PROGRAM Gr01Control
VAR_INPUT
	(* Input variables / Eingang Variablen *)
	bEnable						:BOOL;						(* Enable Gr01Control *)

	(* Instances *)
	fbAxisSawBow				:FB_Gr01SawBow;
	fbAxisAngle					:FB_Gr01Angle;

	fbSawband			 		:FB_Gr01Sawband;

END_VAR
VAR
	(* Enummerations *)

	(* Variables *)
	bAllAxisCtrlEnabled				:BOOL;						(* All axis have controller enabled *)
	bAllAxisStandStill				:BOOL;						(* All axis stand still *)
	bAllAxisNotMoving				:BOOL;						(* All axis not moving *)
	bAllAxisReferenced				:BOOL;						(* All axis referenced *)
	
	BandDistance_m					:LREAL;
	rMachineSawbandSpeed_mmin		:LREAL;

	(* References *)

	(* Interfaces *)

	(* Instances *)
	fbAlarm						:FB_Gr01Alarm;
	fbSafety					:FB_Gr01Safety;
	fbSignals					:FB_Gr01Signals;
	fbUtility					:FB_Gr01Utility;
	rtBtnStart					:R_TRIG;
	
	SawbandVelo					:FB_PosVeloEnc;
	fbLowPassFilter				:FB_LowPassFilter;
	tonSawBandVeloErr			:TON;
	tonSawBandInVelo			:TON;
	TimerVelo					:TON;

END_VAR
VAR CONSTANT
	nFatalErrorMaxIdx			:INT := 0;						(* Maximal index of  using alarms *)
	nErrorMaxIdx				:INT := 19;					(* Maximal index of  using alarms *)
	nWarningMaxIdx				:INT := 0;						(* Maximal index of  using alarms *)
	nMessageMaxIdx				:INT := 1;						(* Maximal index of  using alarms *)
	nHintMaxIdx					:INT := 0;						(* Maximal index of  using alarms *)

	dnFatalErrorBaseIdentNo		:DINT := 11000;				(* Fatal error identification number *)
	dnErrorBaseIdentNo			:DINT := 11100;				(* Error identification number *)
	dnWarningBaseIdentNo		:DINT := 11200;				(* Warning identification number *)
	dnMessageBaseIdentNo		:DINT := 11300;				(* Message identification number *)
	dnHintBaseIdentNo			:DINT := 11400;				(* Hint identification number *)
END_VAR

IF NOT bEnable
THEN
	RETURN;
END_IF;

A_Utility();
A_Safety();
A_Axis();
A_Sawband();
A_Signals();
A_Alarm();

ACTION A_Alarm:

(* Collect and execute input alarms *)
fbAlarm.stAlarmIn.arbError[0].bActive := NOT binGr01LightCurtainOK
                                                		      AND (Gr01Home.fbProcedure.bBusy
                                                      				OR Gr01Auto.fbProcedure.bBusy);
fbAlarm.stAlarmIn.arbError[0].dnCode := dnErrorBaseIdentNo + 0;

fbAlarm.stAlarmIn.arbError[1].bActive := NOT binGr01SawbandRelease
								    AND bgGr00ModeAutomatic
								    AND bgGr00MachineRunning;
fbAlarm.stAlarmIn.arbError[1].dnCode := dnErrorBaseIdentNo + 1;

fbAlarm.stAlarmIn.arbError[2].bActive := FALSE;
fbAlarm.stAlarmIn.arbError[2].dnCode := dnErrorBaseIdentNo + 2;

fbAlarm.stAlarmIn.arbError[3].bActive := FALSE;
fbAlarm.stAlarmIn.arbError[3].dnCode := dnErrorBaseIdentNo + 3;

fbAlarm.stAlarmIn.arbError[4].bActive := fbAxisSawBow.bErrorTerminal;
fbAlarm.stAlarmIn.arbError[4].dnCode := dnErrorBaseIdentNo + 4;

fbAlarm.stAlarmIn.arbError[5].bActive := fbAxisSawBow.fbController.bErrorInit;
fbAlarm.stAlarmIn.arbError[5].dnCode := dnErrorBaseIdentNo + 5;

fbAlarm.stAlarmIn.arbError[6].bActive := fbAxisSawBow.bErrorCtrlEnabled;
fbAlarm.stAlarmIn.arbError[6].dnCode := dnErrorBaseIdentNo + 6;

fbAlarm.stAlarmIn.arbError[7].bActive := fbAxisSawBow.fbController.bError OR fbAxisSawBow.fbMoveManual.bError OR fbAxisSawBow.fbMoveAuto.bError;
fbAlarm.stAlarmIn.arbError[7].dnCode := dnErrorBaseIdentNo + 7;

fbAlarm.stAlarmIn.arbError[8].bActive := fbAxisAngle.bErrorTerminal;
fbAlarm.stAlarmIn.arbError[8].dnCode := dnErrorBaseIdentNo + 8;

fbAlarm.stAlarmIn.arbError[9].bActive := fbAxisAngle.fbController.bErrorInit;
fbAlarm.stAlarmIn.arbError[9].dnCode := dnErrorBaseIdentNo + 9;

fbAlarm.stAlarmIn.arbError[10].bActive := fbAxisAngle.bErrorCtrlEnabled;
fbAlarm.stAlarmIn.arbError[10].dnCode := dnErrorBaseIdentNo + 10;

fbAlarm.stAlarmIn.arbError[11].bActive := fbAxisAngle.fbController.bError OR fbAxisAngle.fbMoveManual.bError OR fbAxisAngle.fbMoveAuto.bError;
fbAlarm.stAlarmIn.arbError[11].dnCode := dnErrorBaseIdentNo + 11;

fbAlarm.stAlarmIn.arbError[12].bActive := fbSawband.bErrorTerminal;
fbAlarm.stAlarmIn.arbError[12].dnCode := dnErrorBaseIdentNo + 12;

fbAlarm.stAlarmIn.arbError[13].bActive := fbSawband.fbController.bErrorInit;
fbAlarm.stAlarmIn.arbError[13].dnCode := dnErrorBaseIdentNo + 13;

fbAlarm.stAlarmIn.arbError[14].bActive := fbSawband.bErrorCtrlEnabled;
fbAlarm.stAlarmIn.arbError[14].dnCode := dnErrorBaseIdentNo + 14;

fbAlarm.stAlarmIn.arbError[15].bActive := fbSawband.fbController.bError OR fbSawband.fbMoveManual.bError OR fbSawband.fbMoveAuto.bError;
fbAlarm.stAlarmIn.arbError[15].dnCode := dnErrorBaseIdentNo + 15;

fbAlarm.stAlarmIn.arbError[16].bActive := FALSE;
fbAlarm.stAlarmIn.arbError[16].dnCode := dnErrorBaseIdentNo + 16;

fbAlarm.stAlarmIn.arbError[17].bActive := GVL_Gr0100.bgGr01SawbandVeloError_1;
fbAlarm.stAlarmIn.arbError[17].dnCode := dnErrorBaseIdentNo + 17;

fbAlarm.stAlarmIn.arbError[18].bActive := GVL_Gr0100.bgGr01SawbandVeloError_2;
fbAlarm.stAlarmIn.arbError[18].dnCode := dnErrorBaseIdentNo + 18;

fbAlarm.stAlarmIn.arbError[19].bActive := (* bgGr00MachineRunning
							AND fbSawband.bCtrlEnabled
							AND fbSawband.bSpeedReached
							AND *) NOT fbSafety.bPipeNotInCrashArea;  (* 20260219 ES/KG *)

fbAlarm.stAlarmIn.arbError[19].dnCode := dnErrorBaseIdentNo + 19;

fbAlarm.stAlarmIn.arbWarning[0].bActive := fbSawband.bErrorVacuumCleanerNOK;
fbAlarm.stAlarmIn.arbWarning[0].dnCode := dnWarningBaseIdentNo + 0;

fbAlarm.stAlarmIn.arbMessage[0].bActive := NOT binGr01LightCurtainOK
							      AND NOT fbAlarm.stAlarmIn.arbError[0].bActive
							      AND NOT fbAlarm.stAlarmOut.arbError[0].bActive;
fbAlarm.stAlarmIn.arbMessage[0].dnCode := dnMessageBaseIdentNo + 0;

fbAlarm.stAlarmIn.arbMessage[1].bActive := NOT binGr01SawbandRelease;
fbAlarm.stAlarmIn.arbMessage[1].dnCode := dnMessageBaseIdentNo + 1;

(* Execute utility *)
fbAlarm(
	etMachineMode := etgGr00MachineMode,
	etMachineState := etgGr00MachineState,
	bNoEStop := bgGr00NoEmergencyStop,
	bConfirmAlarm := bgGr00ConfirmAlarm,
	dtDateTime := stgGr00DateTime.dtDateTime,
	nFatalErrorMaxIdx := nFatalErrorMaxIdx,
	nErrorMaxIdx := nErrorMaxIdx,
	nWarningMaxIdx := nWarningMaxIdx,
	nMessageMaxIdx := nMessageMaxIdx,
	nHintMaxIdx := nHintMaxIdx,
	bMoveInterrupted := bgGr01MoveInterrupted,
	bHomeCompleted := bgGr01HomeCompleted,
	stAlarmOut => stgGr01Alarm.stControl
);
END_ACTION

ACTION A_Axis:

(* Enable axis saw bow *)
stgGr01HMI.stHMITOPLC.lrAxisSawBowNoRefVelo := 10;

fbAxisSawBow(
	bEnable						:= TRUE,
	etMachineMode				:= etgGr00MachineMode,
	etMachineState				:= etgGr00MachineState,
	bMachineStandstill			:= bgGr00MachineStandstill,
	bNoEStop					:= bgGr00NoEmergencyStop,
	bPowerSupplyOn				:= bgGr00PowerSupplyOk,
	bSafetyOK					:= bgGr01LightCurtainOK
								   AND bgGr00AllDoorsClosedLocked,
	bCtrlInterrupt				:= FALSE,
	bMoveRelease				:= TRUE,
	bPlusRelease				:= TRUE,
	bMinusRelease				:= TRUE,
	bSignalReference			:= NOT binGr01AxisSawBowLimitMax,
	bSignalHWLimitMax			:= NOT binGr01AxisSawBowLimitMax,
	bSignalHWLimitMin			:= NOT binGr01AxisSawBowLimitMin,
	lrSoftLimitMax				:= stgGr01HMI.stHMITOPLC.lrAxisSawBowSoftLimitMax,
	lrSoftLimitMin				:= stgGr01HMI.stHMITOPLC.lrAxisSawBowSoftLimitMin,
	bConfirmAlarm				:= bgGr00ConfirmAlarm,
	bTipPlus					:= stgGr01HMI.stHMITOPLC.bBtnAxisSawBowPlus,
	bTipMinus					:= stgGr01HMI.stHMITOPLC.bBtnAxisSawBowMinus,
	lrManualVelocity			:= stgGr01HMI.stHMITOPLC.lrAxisSawBowManualVelo,
	lrNoRefVelocity				:= stgGr01HMI.stHMITOPLC.lrAxisSawBowNoRefVelo,
	bVelocityLimitEn			:= FALSE,
	lrAcceleration				:= 100.0,
	lrDeceleration				:= 100.0,
	lrJerk						:= 100.0,
	lrOverride					:= fbUtility.rActOverride,
	lrExtOverride				:= 0.0,
	dnRatioNumerator			:= 1,
	udnRatioDenominator			:= 1,
	bEngineTorqueLimitEn		:= FALSE,
	lrEngineTorque				:= 200.0,
	tControllerOff				:= tgGr01ControllerOff,
	bWithAbsoluteEncoder		:= FALSE,
	lrOriginShiftPos			:= stgGr01HMI.stHMITOPLC.lrAxisSawBowOriginShiftPos,
	bVeloForceCtrlEn			:= FALSE,
	tAdsTimeOut					:= DEFAULT_ADS_TIMEOUT,
	bHomeCompleted				:= bgGr01HomeCompleted,
	Drive						:= GVL_Gr01Interface.igGr01DriveSawBow,
	Axis						:= GVL_Gr01Interface.igGr01AxisSawBow,
	MasterAxis					:= GVL_Gr00Interface.iAxisDummy,
	
	lrActPosition				=> stgGr01HMI.stPLCTOHMI.lrAxisSawBowActPos,
	lrActVelocity				=> stgGr01HMI.stPLCTOHMI.lrAxisSawBowActVelo,
	lrActForce					=> stgGr01HMI.stPLCTOHMI.lrAxisSawBowActForce
);

(* Enable Axis angle *)
stgGr01HMI.stHMITOPLC.lrAxisAngleNoRefVelo := 10;



fbAxisAngle(
	bEnable						:= TRUE,

	etMachineMode				:= etgGr00MachineMode,
	etMachineState				:= etgGr00MachineState,
	bMachineStandstill			:= bgGr00MachineStandstill,
	bNoEStop					:= bgGr00NoEmergencyStop,
	bPowerSupplyOn				:= bgGr00PowerSupplyOk,
	bSafetyOK					:= bgGr01LightCurtainOK
								   AND bgGr00AllDoorsClosedLocked,
	bCtrlInterrupt				:= FALSE,
	bMoveRelease				:= TRUE,
	bMoveInterrupt				:= FALSE,
	bPlusRelease				:= TRUE,
	bMinusRelease				:= TRUE,	(*stgGr00HMI.stHMITOPLC.bSafetyInterlockOff*)
	bHWSignalLimitMax			:= NOT binGr01AxisAngleLimitMax,
	bHWSignalLimitMin			:= NOT binGr01AxisAngleLimitMin,
	lrSoftLimitMax				:= stgGr01HMI.stHMITOPLC.lrAxisAngleSoftLimitMax,
	lrSoftLimitMin				:= stgGr01HMI.stHMITOPLC.lrAxisAngleSoftLimitMin,
	bConfirmAlarm				:= bgGr00ConfirmAlarm,
	bTipPlus					:= stgGr01HMI.stHMITOPLC.bBtnAxisAnglePlus,
	bTipMinus					:= stgGr01HMI.stHMITOPLC.bBtnAxisAngleMinus,
	lrManualVelocity			:= stgGr01HMI.stHMITOPLC.lrAxisAngleManualVelo,
	lrVelocityNoRef				:= stgGr01HMI.stHMITOPLC.lrAxisAngleNoRefVelo,
	bVelocityLimitEn			:= FALSE,
	lrAcceleration				:= 100.0,
	lrDeceleration				:= 100.0,
	lrJerk						:= 100.0,
	lrOverride					:= fbUtility.rActOverride,
	bEngineTorqueLimitEn		:= FALSE,
	lrEngineTorque				:= 200.0,
	tControllerOff				:= tgGr01ControllerOff,
	lrScalingNum				:= lrgGr01AxisAnglePath,
	udnScalingDenom				:= udngGr01AxisAngleInc,
	bWithAbsoluteEncoder		:= TRUE,
	udnIncEnc					:= udninGr01IncAxisAngle,
	lrOriginShift				:= stgGr01HMI.stHMITOPLC.lrAxisAngleOriginShiftPos,
	lrTaskCycle					:= lrgActCycleTime,
	tAdsTimeOut					:= DEFAULT_ADS_TIMEOUT,
	bHomeCompleted				:= bgGr01HomeCompleted,
	Drive						:= GVL_Gr01Interface.igGr01DriveSawAngle,
	Axis						:= GVL_Gr01Interface.igGr01AxisSawAngle,
	MasterAxis					:= GVL_Gr00Interface.iAxisDummy,
	
	lrActPosition				=> stgGr01HMI.stPLCTOHMI.lrAxisAngleActPos,
	lrActVelocity				=> stgGr01HMI.stPLCTOHMI.lrAxisAngleActVelo
);
END_ACTION

ACTION A_Safety:

(* Execute safety *)
fbSafety(
	bLightCurtain := binGr01LightCurtainOK,
	bConfirmLightCurtain := (bgGr00ConfirmAlarm
			                            OR etgGr00MachineMode = ET_MachineMode_eManual
			                            OR etgGr00MachineMode = ET_MachineMode_eHome
			                            OR etgGr00MachineMode = ET_MachineMode_eAutomatic
			                            OR stgGr00HMI.stHMITOPLC.bSafetyInterlockOff)
					         AND NOT stgGr01Alarm.stControl.arbError[0].bActive,
	tLightCurtainDelay := tgGr01LightCurtainDelay,
	bLightCurtainOK => bgGr01LightCurtainOK,
	bConfirmedLightCurtain => boutGr01ConfLightCurtain,
	bNotInCrashArea => bgGr01NotInCrashArea
);

bgGr01SafetyActive := fbAxisSawBow.bSafetyLock
				        OR fbAxisAngle.bSafetyLock;
END_ACTION

ACTION A_Sawband:

fbSawband(
	bEnable						:= TRUE,
	bOccupied					:= FALSE,
	etMachineMode				:= etgGr00MachineMode,
	etMachineState				:= etgGr00MachineState,
	bMachineStandstill			:= bgGr00MachineStandstill,
	bNoEStop					:= bgGr00NoEmergencyStop,
	bPowerSupplyOn				:= bgGr00PowerSupplyOk,	//fbStoeberPS6A34.bOn, // Keine Eingänge vorhanden
	bSafetyOK					:= bgGr01LightCurtainOK								   AND bgGr00AllDoorsClosedLocked,
	bSafetyDriveEnabled			:= TRUE,
	bCtrlInterrupt				:= FALSE,
	bMoveRelease				:= TRUE,
	bPlusRelease				:= TRUE,
	bMinusRelease				:= FALSE,
	bSignalReference			:= FALSE,
	bSignalHWLimitMax			:= FALSE,
	bSignalHWLimitMin			:= FALSE,
	lrSoftLimitMax				:= 0,
	lrSoftLimitMin				:= 0,
	etHomingMode				:= MC_DefaultHoming,
	bConfirmAlarm				:= bgGr00ConfirmAlarm,
	bTipPlus					:= stgGr01HMI.stHMITOPLC.bBtnSawbandPlus,
	bTipMinus					:= False,
	lrTipDistance				:= 0,
	lrManualVelocity			:= stgGr01HMI.stHMITOPLC.rSawbandManualSpeed / 3.28084,
	lrAutoVelocity				:= stgGr01HMI.stHMITOPLC.rSawbandAutoSpeed / 3.28084,
	lrNoRefVelocity				:= 30,
	bVelocityLimitEn			:= FALSE,
	lrAcceleration				:= 5000,
	lrDeceleration				:= 5000,
	lrJerk						:= 30000,
	lrOverride					:= 100.0,
	bExtOverrideEn				:= FALSE,
	dnRatioNumerator			:= 1,
	udnRatioDenominator			:= 1,
	bEngineTorqueLimitEn		:= FALSE,
	lrEngineTorque				:= 400,
	bPosLagMonitoringEn			:= FALSE,
	tControllerOff				:= tgGr01ControllerOff,
	bWithAbsoluteEncoder		:= FALSE,
	bVeloForceCtrlEn			:= FALSE,
	tAdsTimeOut					:= DEFAULT_ADS_TIMEOUT,
	bHomeCompleted				:= bgGr01HomeCompleted,
	Drive						:= GVL_Gr01Interface.igGr01DriveSawBand,
	Axis						:= GVL_Gr01Interface.igGr01AxisSawBand,
	MasterAxis					:= GVL_Gr00Interface.iAxisDummy,

	lrActVelocity				=> GVL_Gr01HMI.stgGr01HMI.stPLCTOHMI.lrSawbandActSpeed,
	bSawbandAirOn 				=> boutGr01SawbandAirOn
);

rMachineSawbandSpeed_mmin := stgGr01HMI.stHMITOPLC.rSawbandAutoSpeed / 3.28084;

////////////// Sawband Velo Scaling

SawbandVelo(
	bEnable				:= TRUE , 
	dwEncCurrentValue	:= GVL_GR01IO.udninGr01CounterSawbandSpeed, 
	udnScalingDenom		:= uiImpulsDiscAmount , 	
	lrScalingNum		:= rRaddurchmesser_mm*PI, 	
	tCycleTime			:= GVL_Gr00Init.tPLC_TaskCycleTime_ms, 					
	lrCurrentPos		=> , 
	lrCurrentVelo		=> ,			(* [mm/ms] same as [m/s]*)
);
	
BandDistance_m := SawbandVelo.lrCurrentPos / 1000;
GVL_Gr01Init.lrgGr01SawingSpeed := SawbandVelo.lrCurrentVelo * 60;		(* [m/min] *)

	fbLowPassFilter(
	bEnable			:= TRUE , 
	lrIn			:= GVL_Gr01Init.lrgGr01SawingSpeed, 
	lrKp			:= 1, 
	tT1				:= T#600MS , 
	tCycletime		:= GVL_Gr00Init.tPLC_TaskCycleTime_ms, 
	lrOut			=> GVL_Gr01Init.lrgGr01SawingSpeed

);
//////////////
GVL_Gr01HMI.stgGr01HMI.stHMITOPLC.rSawbandAutoSpeed := GVL_Gr01Init.lrgGr01SawingSpeed;
	
	
////////////// Sawband Velo Error -> never reaches target speed
tonSawBandInVelo(
					IN:= NOT GVL_GR0100.bgGr01SawbandVeloError_1 AND (ABS(GVL_Gr01Interface.igGr01AxisSawBand.NcToPlc.ActVelo) - ABS(GVL_Gr01Interface.igGr01AxisSawBand.NcToPlc.SetVelo)< 100),
					PT := T#3S);
					
GVL_GR0100.bgGr01SawbandInSpeed := GVL_Gr01Init.lrgGr01SawingSpeed > (rMachineSawbandSpeed_mmin * 0.8 * fbSawband.lrOverride/100)
							AND (tonSawBandInVelo.Q OR GVL_Gr01HMI.stgGr01HMI.stHMITOPLC.bBtnSawbandPlus);
							
TimerVelo(
	IN:= NOT GVL_GR0100.bgGr01SawbandInSpeed AND NOT GVL_GR0100.bgGr01SawbandVeloError_1 AND GVL_Gr0000.bgGr00NoEmergencyStop, 
	PT:=T#10S
		); 
		
GVL_GR0100.bgGr01SawbandVeloError_1 := TimerVelo.Q; 


//Sawband velocity error -> lost target speed
tonSawBandVeloErr(
					IN:=ABS(GVL_Gr01Interface.igGr01AxisSawBand.NcToPlc.ActVelo) < ABS(GVL_Gr01Interface.igGr01AxisSawBand.NcToPlc.SetVelo *0.8),
					PT := T#500MS);

GVL_GR0100.bgGr01SawbandVeloError_2 := tonSawBandInVelo.Q;



(* Old FB)
(* Enable sawband *)
fbSawband(
	bEnable := TRUE,
	lrScalingNum := lrgGr01SawbandDistance,
	udnScalingDenom := udngGr01SawbandInc,
	etMachineMode := etgGr00MachineMode,
	etMachineState := etgGr00MachineState,
	bNoEStop := bgGr00NoEmergencyStop,
	bPowerSupplyOn := bgGr00PowerSupplyOk,
	bSafetyOK := bgGr01LightCurtainOK
			        AND bgGr00AllDoorsClosedLocked,
	bAirPressureOK := bgGr00AirPressureOK,
	bMachineStandstill := bgGr00MachineStandstill,
	bCtrlInterrupt := FALSE,
	bMoveRelease := TRUE,
	bMoveInterrupt := FALSE,
	bTipPlus := stgGr01HMI.stHMITOPLC.bBtnSawbandPlus,
	bTipMinus := FALSE(*stgGr01HMI.stHMITOPLC.bBtnSawbandMinus*),
	bPlusRelease := TRUE,
	bMinusRelease := TRUE,
	bHandSawbandAirOn := stgGr01HMI.stHMITOPLC.bBtnSawbandAirOn,
	bHandVacuumCleanerOn := stgGr01HMI.stHMITOPLC.bBtnVacuumCleanerOn,
	bExtOverrideEn := FALSE,
	lrManualSpeed := stgGr01HMI.stHMITOPLC.rSawbandManualSpeed / 3.28084,
	lrAutoSpeed := stgGr01HMI.stHMITOPLC.rSawbandAutoSpeed  / 3.28084,
	bSpeedLimitEn := TRUE,
	lrSpeedMin := 0, (* m/min *)
	lrSpeedMax := 400, (* m/min  SY 650*)
	lrAcceleration := 100.0,
	lrDeceleration := 100.0,
	lrJerk := 100.0,
	bEngineTorqueLimitEn := FALSE,
	lrEngineTorque := 200.0,
	bSawbandMotorNOK := binGr01SawbandMotorNOK,
	bSawbandBroken := NOT binGr01SawbandNoBroken,
	bVacuumCleanerMotorNOK := binGr01VacuumCleanerMotorNOK,
	udnIncEnc := udninGr01CounterSawbandSpeed,
	lrTaskCycle := lrgActCycleTime,
	bConfirmAlarm := bgGr00ConfirmAlarm,
	tSawbandAirOffDelay := tgGr01SawbandAirOffDelay,
	tVacuumCleanerOffDelay := tgGr01VacuumCleanerOffDelay,
	tSawbandReadyDelay := tgGr01SawbandReadyDelay,
	tSpeedNoConstant := tgGr01SpeedNoConstant,
	tControllerOff := tgGr01ControllerOff,
	tAdsTimeOut := DEFAULT_ADS_TIMEOUT,
	bHomeCompleted := bgGr01HomeCompleted,
	Drive := igGr01DriveSawband,
	Axis := igGr01AxisSawband,
	lrActSpeed => stgGr01HMI.stPLCTOHMI.lrSawbandActSpeed,
	bSawbandAirOn => boutGr01SawbandAirOn,
	bVacuumCleanerOn => boutGr01VacuumCleanerOn
);
*)
END_ACTION

ACTION A_Signals:

(* Execute signals *)
fbSignals(
	etMachineMode := etgGr00MachineMode,
	etMachineState := etgGr00MachineState,
	bMachineRunning := bgGr00MachineRunning,
	bExecutedProcess := fbUtility.arbExeProcess[1]
					      OR fbUtility.arbExeProcess[2]
					      OR fbUtility.arbExeProcess[3],
	stBlinker := stgGr00Blinker,
	bBulbBtnStart => boutGr01BulbBtnStart,
	bBulbBtnStop => boutGr01BulbBtnStop,
);

(* Detect all axis controller enabled *)
bAllAxisCtrlEnabled := F_ChkAllAxisEnabled(
	bEnable := TRUE,
	bEnabledAxis1 := Gr01Control.fbAxisSawBow.bCtrlEnabled,
	bEnabledAxis2 := Gr01Control.fbAxisAngle.bCtrlEnabled,
	bEnabledAxis3 := TRUE,
	bEnabledAxis4 := TRUE,
	bEnabledAxis5 := TRUE,
	bEnabledAxis6 := TRUE,
	bEnabledAxis7 := TRUE,
	bEnabledAxis8 := TRUE,
	bEnabledAxis9 := TRUE,
	bEnabledAxis10 := TRUE
);

(* Detect all axis stand still *)
bAllAxisStandStill := F_ChkAllAxisStandStill(
	bEnable := TRUE,
	bAxis1StandStill := Gr01Control.fbAxisSawBow.bStandStill, 		// igGr01AxisSawBow.stAxisStatus.bStandStill,
	bAxis2StandStill := Gr01Control.fbAxisAngle.bStandStill,		// igGr01AxisAngle.stAxisStatus.bStandStill,
	bAxis3StandStill := TRUE,
	bAxis4StandStill := TRUE,
	bAxis5StandStill := TRUE,
	bAxis6StandStill := TRUE,
	bAxis7StandStill := TRUE,
	bAxis8StandStill := TRUE,
	bAxis9StandStill := TRUE,
	bAxis10StandStill := TRUE,
);

(* Detect all axis not moving *)
bAllAxisNotMoving := F_ChkAllAxisNotMoving(
	bEnable := TRUE,
	bAxis1NotMoving := Gr01Control.fbAxisSawBow.bNotMoving, 		
	bAxis2NotMoving := Gr01Control.fbAxisAngle.bNotMoving,
	bAxis3NotMoving := TRUE,
	bAxis4NotMoving := TRUE,
	bAxis5NotMoving := TRUE,
	bAxis6NotMoving := TRUE,
	bAxis7NotMoving := TRUE,
	bAxis8NotMoving := TRUE,
	bAxis9NotMoving := TRUE,
	bAxis10NotMoving := TRUE
);

(* Detect all axis referenced *)
bAllAxisReferenced := F_ChkAllAxisReferenced(
	bEnable := TRUE,
	bReferencedAxis1 := Gr01Control.fbAxisSawBow.bReferenced,
	bReferencedAxis2 := Gr01Control.fbAxisAngle.bReferenced,
	bReferencedAxis3 := TRUE,
	bReferencedAxis4 := TRUE,
	bReferencedAxis5 := TRUE,
	bReferencedAxis6 := TRUE,
	bReferencedAxis7 := TRUE,
	bReferencedAxis8 := TRUE,
	bReferencedAxis9 := TRUE,
	bReferencedAxis10 := TRUE
);
END_ACTION

ACTION A_Utility:

(* Execute utility *)

(* Start program *)
rtBtnStart(CLK := binGr00PushBtnStart OR stgGr00HMI.stHMITOPLC.bBtnStart);

fbUtility.arbStartProcess[1] := rtBtnStart.Q
						 AND etgGr00MachineState = ET_MachineState_eAutoExe;
fbUtility.arbStopProcess[1] := etgGr00MachineState <> ET_MachineState_eAutoExe;
fbUtility.arbSteppingProcess[1] := stgGr01HMI.stHMITOPLC.bBtnSteppingProcess;
arbgGr01StartProcess[1] := fbUtility.arbExeProcess[1];

fbUtility(
	etMachineMode := etgGr00MachineMode,
	etMachineState := etgGr00MachineState,
	bAutoCompleted := bgGr00AutoCompleted
					  AND bgGr01AutoCompleted
					  AND bgGr02AutoCompleted
					  AND bgGr05AutoCompleted
					  AND bgGr00MachineStandstill
					  AND etgGr00MachineState <> ET_MachineState_eAutoExe,
	bHomeCompleted := bgGr01HomeCompleted,
	bExeCounter := bgGr01AutoCompleted,
	bLaserOnOff := stgGr01HMI.stHMITOPLC.bBtnLaserOn,
	bStartTime := Gr01Control.fbUtility.arbStartProcess[1]
				OR Gr01Control.fbUtility.arbStartProcess[2]
				OR Gr01Control.fbUtility.arbStopProcess[3],
	bStopTime := bgGr01AutoCompleted
				OR fbUtility.arbStopProcess[1]
				OR fbUtility.arbStopProcess[2]
				OR fbUtility.arbStopProcess[3],
	bLifetimeOn := NOT fbSawband.bNotMoving,
	bResetLifetimeAll := FALSE,
	bResetLifetime := stgGr01HMI.stHMITOPLC.bResetLifetime,
	sLifetimeFilePath := sgGr01LifetimeFilePath,
	sLifetimeFileName := sgGr01LifetimeFileName,
	bPipeIdentify := NOT binGr01PipeNoIdentify,
	rGlobalOverride := rgGr00Override,
	rLocalOverride := stgGr01HMI.stHMITOPLC.rOverride,
	lrLifetimeAll => stgGr01HMI.stPLCTOHMI.lrLifetime,
	lrLifetimeAfterReset => stgGr01HMI.stPLCTOHMI.lrLifetimeAfterReset,
	lrLifetimeAfterTrunOn => stgGr01HMI.stPLCTOHMI.lrLifetimeAfterTurnOn,
	udnCounterTotal := stgGr01HMI.stPLCTOHMI.udnCounterTotal,
	bLaserOn => boutGr01LaserOn,
	bPipePresent => bgGr01PipePresent
);
END_ACTION

END_PROGRAM

(* stored: Version 1.1.0.1, ProductVersion 3.1.4024.15
   POU Gr01Control: Id {2dac79ca-e47b-4d2d-839b-3f84db7e801e}, SpecialFunc None
   Action A_Alarm: Id {e9f90f32-b3c1-41b6-ad3f-b8525a491730}
   Action A_Axis: Id {e1fcb53e-2fd3-4612-85cf-3d8298151cc6}
   Action A_Safety: Id {fb2b49ed-022e-4de4-a5f8-c1ee5bdd8a09}
   Action A_Sawband: Id {96a1aa51-3ac5-4b37-a51d-5bd0b216fe25}
   Action A_Signals: Id {970ec869-7b46-429c-a071-32fe1da01a64}
   Action A_Utility: Id {a99fa86f-8295-4f3e-9137-945607a2d57f} *)
